Fanuc KAREL source: KB00033.KL

PROGRAM KB00033
%NOLOCKGROUP
%ENVIRONMENT STRNG
VAR
  P1: CONFIG
  P2: STRING[80]
  P3: INTEGER
BEGIN
  P2 = 'A'
  P3 = 1
  CNV_CNF_STRG(P1, P2, P3)
END KB00033
